# EPICS autosave request: iocs/meascomp/db/measCompMCS_settings.req
$(P)PresetReal
$(P)Dwell
$(P)Prescale
$(P)ChannelAdvance
$(P)MCSCounter1Enable
$(P)MCSCounter2Enable
$(P)MCSCounter3Enable
$(P)MCSCounter4Enable
$(P)MCSCounter5Enable
$(P)MCSCounter6Enable
$(P)MCSCounter7Enable
$(P)MCSCounter8Enable
$(P)MCSDIOEnable
$(P)PrescaleCounter
$(P)Point0Action
$(P)ReadAll.SCAN
$(P)NuseAll
$(P)EnableClientWait
$(P)TrigMode
